FUNCTION_BLOCK FB_Valve
VAR_OUTPUT
	bOpen AT %Q* : BOOL;   // solenoid
END_VAR
VAR
	tOpened : TIME;
END_VAR

;

METHOD Open
bOpen := TRUE;
END_METHOD

PROPERTY IsOpen : BOOL
GET
IsOpen := bOpen;
END_GET
END_PROPERTY

END_FUNCTION_BLOCK

(* stored: Version 1.1.0.1, ProductVersion 3.1.4024.12
   POU FB_Valve: Id {aaaaaaaa-0000-0000-0000-000000000004}, SpecialFunc None
   Method Open: Id {aaaaaaaa-0000-0000-0000-000000000005}
   Property IsOpen: Id {aaaaaaaa-0000-0000-0000-000000000006}
   Get Get: Id {aaaaaaaa-0000-0000-0000-000000000007} *)
